// TIA Portal V20 export
FUNCTION_BLOCK "FB_LD_PressDemoAuto"   // FB, LAD
{ S7_Optimized_Access := 'TRUE' }
// stored: AutoNumber true
   VAR_INPUT
      Run { ExternalWritable := 'False'} : Bool;
      Reset { ExternalWritable := 'False'} : Bool;
      OwnerIndex { ExternalWritable := 'False'} : DInt;
      Delta { ExternalWritable := 'False'} : Time;
      TransferSettleTime { ExternalWritable := 'False'} : Time;
      PartQuality { ExternalWritable := 'False'} : Bool;
      RequireTwoHandStart { ExternalWritable := 'False'} : Bool;
      SourcePath { ExternalWritable := 'False'} : String[80];
      PartPresent { ExternalWritable := 'False'} : Bool;
      AirPressureOk { ExternalWritable := 'False'} : Bool;
      TwoHandHeld { ExternalWritable := 'False'} : Bool;
      StartPulse { ExternalWritable := 'False'} : Bool;
      PressSettleTime { ExternalWritable := 'False'} : Time;
   END_VAR
   VAR_IN_OUT
      PressRam { ExternalAccessible := 'False'; ExternalVisible := 'False'; ExternalWritable := 'False'} : "FB_CylinderCM";
      Door { ExternalAccessible := 'False'; ExternalVisible := 'False'; ExternalWritable := 'False'} : "FB_CylinderCM";
      PartSlide { ExternalAccessible := 'False'; ExternalVisible := 'False'; ExternalWritable := 'False'} : "FB_CylinderCM";
      Core { ExternalAccessible := 'False'; ExternalVisible := 'False'; ExternalWritable := 'False'} : "FRK_Core";
      Unit { ExternalAccessible := 'False'; ExternalVisible := 'False'; ExternalWritable := 'False'} : "FRK_Unit";
      Status { ExternalAccessible := 'False'; ExternalVisible := 'False'; ExternalWritable := 'False'} : "ST_ModuleStatus";
      Part { ExternalAccessible := 'False'; ExternalVisible := 'False'; ExternalWritable := 'False'} : "ST_PartContext";
      AlarmLog { ExternalAccessible := 'False'; ExternalVisible := 'False'; ExternalWritable := 'False'} : "FRK_AlarmLog";
   END_VAR
   VAR
      Seq { ExternalWritable := 'False'} : "FRK_SequenceCtx";
      Row1 { ExternalWritable := 'False'} : "FRK_SequenceRow";
      Row2 { ExternalWritable := 'False'} : "FRK_SequenceRow";
      Row3 { ExternalWritable := 'False'} : "FRK_SequenceRow";
      Row4 { ExternalWritable := 'False'} : "FRK_SequenceRow";
      Row5 { ExternalWritable := 'False'} : "FRK_SequenceRow";
      Row6 { ExternalWritable := 'False'} : "FRK_SequenceRow";
      Row7 { ExternalWritable := 'False'} : "FRK_SequenceRow";
      Row8 { ExternalWritable := 'False'} : "FRK_SequenceRow";
      Row9 { ExternalWritable := 'False'} : "FRK_SequenceRow";
      Row10 { ExternalWritable := 'False'} : "FRK_SequenceRow";
      Row11 { ExternalWritable := 'False'} : "FRK_SequenceRow";
      Row12 { ExternalWritable := 'False'} : "FRK_SequenceRow";
      Row13 { ExternalWritable := 'False'} : "FRK_SequenceRow";
      Row14 { ExternalWritable := 'False'} : "FRK_SequenceRow";
      Row15 { ExternalWritable := 'False'} : "FRK_SequenceRow";
      Row16 { ExternalWritable := 'False'} : "FRK_SequenceRow";
      At0 { ExternalAccessible := 'False'; ExternalVisible := 'False'; ExternalWritable := 'False'} : Bool;
      At100 { ExternalAccessible := 'False'; ExternalVisible := 'False'; ExternalWritable := 'False'} : Bool;
      At110 { ExternalAccessible := 'False'; ExternalVisible := 'False'; ExternalWritable := 'False'} : Bool;
      At130 { ExternalAccessible := 'False'; ExternalVisible := 'False'; ExternalWritable := 'False'} : Bool;
      At150 { ExternalAccessible := 'False'; ExternalVisible := 'False'; ExternalWritable := 'False'} : Bool;
      At170 { ExternalAccessible := 'False'; ExternalVisible := 'False'; ExternalWritable := 'False'} : Bool;
      At180 { ExternalAccessible := 'False'; ExternalVisible := 'False'; ExternalWritable := 'False'} : Bool;
      At185 { ExternalAccessible := 'False'; ExternalVisible := 'False'; ExternalWritable := 'False'} : Bool;
      At190 { ExternalAccessible := 'False'; ExternalVisible := 'False'; ExternalWritable := 'False'} : Bool;
      At200 { ExternalAccessible := 'False'; ExternalVisible := 'False'; ExternalWritable := 'False'} : Bool;
      At210 { ExternalAccessible := 'False'; ExternalVisible := 'False'; ExternalWritable := 'False'} : Bool;
      At215 { ExternalAccessible := 'False'; ExternalVisible := 'False'; ExternalWritable := 'False'} : Bool;
      At220 { ExternalAccessible := 'False'; ExternalVisible := 'False'; ExternalWritable := 'False'} : Bool;
      At230 { ExternalAccessible := 'False'; ExternalVisible := 'False'; ExternalWritable := 'False'} : Bool;
      At240 { ExternalAccessible := 'False'; ExternalVisible := 'False'; ExternalWritable := 'False'} : Bool;
      At999 { ExternalAccessible := 'False'; ExternalVisible := 'False'; ExternalWritable := 'False'} : Bool;
      Ready1 { ExternalAccessible := 'False'; ExternalVisible := 'False'; ExternalWritable := 'False'} : Bool;
      Ready2 { ExternalAccessible := 'False'; ExternalVisible := 'False'; ExternalWritable := 'False'} : Bool;
      Ready3 { ExternalAccessible := 'False'; ExternalVisible := 'False'; ExternalWritable := 'False'} : Bool;
      Ready4 { ExternalAccessible := 'False'; ExternalVisible := 'False'; ExternalWritable := 'False'} : Bool;
      Ready5 { ExternalAccessible := 'False'; ExternalVisible := 'False'; ExternalWritable := 'False'} : Bool;
      Advance { ExternalAccessible := 'False'; ExternalVisible := 'False'; ExternalWritable := 'False'} : Bool;
      Cycle { ExternalAccessible := 'False'; ExternalVisible := 'False'; ExternalWritable := 'False'} : "ST_PressDemoCycle";
      LoadPosition { ExternalAccessible := 'False'; ExternalVisible := 'False'; ExternalWritable := 'False'} : "FB_PressDemoLoadPosition";
      LoadDone { ExternalAccessible := 'False'; ExternalVisible := 'False'; ExternalWritable := 'False'} : Bool;
      LoadActive { ExternalAccessible := 'False'; ExternalVisible := 'False'; ExternalWritable := 'False'} : Bool;
   END_VAR
BEGIN

REGION Network 1
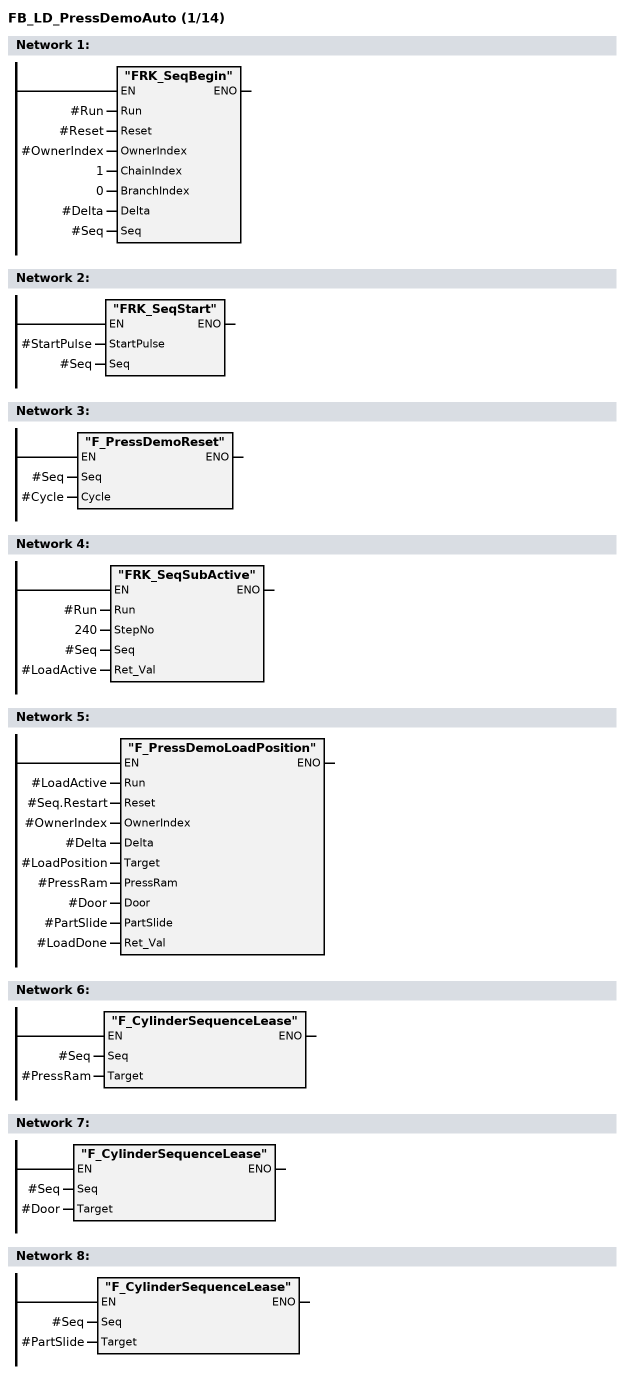
   RUNG wire#powerrail
      "FRK_SeqBegin"(Run := #Run, Reset := #Reset, OwnerIndex := #OwnerIndex, ChainIndex := 1, BranchIndex := 0, Delta := #Delta, Seq := #Seq)
   END_RUNG
   // the same network as SCL:
   "FRK_SeqBegin"(Run := #Run,
                  Reset := #Reset,
                  OwnerIndex := #OwnerIndex,
                  ChainIndex := 1,
                  BranchIndex := 0,
                  Delta := #Delta,
                  Seq := #Seq);
END_REGION

REGION Network 2
   RUNG wire#powerrail
      "FRK_SeqStart"(StartPulse := #StartPulse, Seq := #Seq)
   END_RUNG
   // the same network as SCL:
   "FRK_SeqStart"(StartPulse := #StartPulse, Seq := #Seq);
END_REGION

REGION Network 3
   RUNG wire#powerrail
      "F_PressDemoReset"(Seq := #Seq, Cycle := #Cycle)
   END_RUNG
   // the same network as SCL:
   "F_PressDemoReset"(Seq := #Seq, Cycle := #Cycle);
END_REGION

REGION Network 4
   RUNG wire#powerrail
      "FRK_SeqSubActive"(Run := #Run, StepNo := 240, Seq := #Seq, Ret_Val := #LoadActive)
   END_RUNG
   // the same network as SCL:
   "FRK_SeqSubActive"(Run := #Run, StepNo := 240, Seq := #Seq, Ret_Val := #LoadActive);
END_REGION

REGION Network 5
   RUNG wire#powerrail
      "F_PressDemoLoadPosition"(Run := #LoadActive, Reset := #Seq.Restart, OwnerIndex := #OwnerIndex, Delta := #Delta, Target := #LoadPosition, PressRam := #PressRam, Door := #Door, PartSlide := #PartSlide, Ret_Val := #LoadDone)
   END_RUNG
   // the same network as SCL:
   "F_PressDemoLoadPosition"(Run := #LoadActive,
                           Reset := #Seq.Restart,
                           OwnerIndex := #OwnerIndex,
                           Delta := #Delta,
                           Target := #LoadPosition,
                           PressRam := #PressRam,
                           Door := #Door,
                           PartSlide := #PartSlide,
                           Ret_Val := #LoadDone);
END_REGION

REGION Network 6
   RUNG wire#powerrail
      "F_CylinderSequenceLease"(Seq := #Seq, Target := #PressRam)
   END_RUNG
   // the same network as SCL:
   "F_CylinderSequenceLease"(Seq := #Seq, Target := #PressRam);
END_REGION

REGION Network 7
   RUNG wire#powerrail
      "F_CylinderSequenceLease"(Seq := #Seq, Target := #Door)
   END_RUNG
   // the same network as SCL:
   "F_CylinderSequenceLease"(Seq := #Seq, Target := #Door);
END_REGION

REGION Network 8
   RUNG wire#powerrail
      "F_CylinderSequenceLease"(Seq := #Seq, Target := #PartSlide)
   END_RUNG
   // the same network as SCL:
   "F_CylinderSequenceLease"(Seq := #Seq, Target := #PartSlide);
END_REGION

REGION Network 9
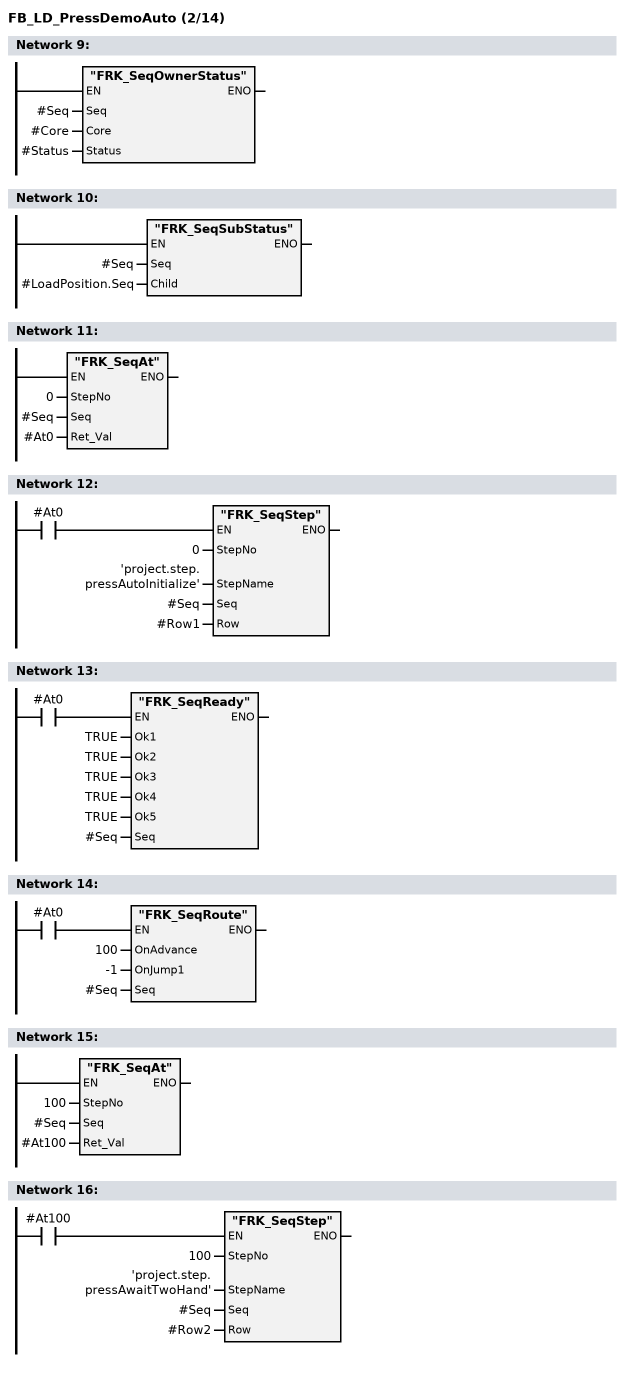
   RUNG wire#powerrail
      "FRK_SeqOwnerStatus"(Seq := #Seq, Core := #Core, Status := #Status)
   END_RUNG
   // the same network as SCL:
   "FRK_SeqOwnerStatus"(Seq := #Seq, Core := #Core, Status := #Status);
END_REGION

REGION Network 10
   RUNG wire#powerrail
      "FRK_SeqSubStatus"(Seq := #Seq, Child := #LoadPosition.Seq)
   END_RUNG
   // the same network as SCL:
   "FRK_SeqSubStatus"(Seq := #Seq, Child := #LoadPosition.Seq);
END_REGION

REGION Network 11
   RUNG wire#powerrail
      "FRK_SeqAt"(StepNo := 0, Seq := #Seq, Ret_Val := #At0)
   END_RUNG
   // the same network as SCL:
   "FRK_SeqAt"(StepNo := 0, Seq := #Seq, Ret_Val := #At0);
END_REGION

REGION Network 12
   IF #At0 THEN
       "FRK_SeqStep"(StepNo := 0, StepName := 'project.step.pressAutoInitialize', Seq := #Seq, Row := #Row1);
   END_IF;
END_REGION

REGION Network 13
   IF #At0 THEN
       "FRK_SeqReady"(Ok1 := TRUE, Ok2 := TRUE, Ok3 := TRUE, Ok4 := TRUE, Ok5 := TRUE, Seq := #Seq);
   END_IF;
END_REGION

REGION Network 14
   IF #At0 THEN "FRK_SeqRoute"(OnAdvance := 100, OnJump1 := -1, Seq := #Seq); END_IF;
END_REGION

REGION Network 15
   RUNG wire#powerrail
      "FRK_SeqAt"(StepNo := 100, Seq := #Seq, Ret_Val := #At100)
   END_RUNG
   // the same network as SCL:
   "FRK_SeqAt"(StepNo := 100, Seq := #Seq, Ret_Val := #At100);
END_REGION

REGION Network 16
   IF #At100 THEN
       "FRK_SeqStep"(StepNo := 100, StepName := 'project.step.pressAwaitTwoHand', Seq := #Seq, Row := #Row2);
   END_IF;
END_REGION

REGION Network 17
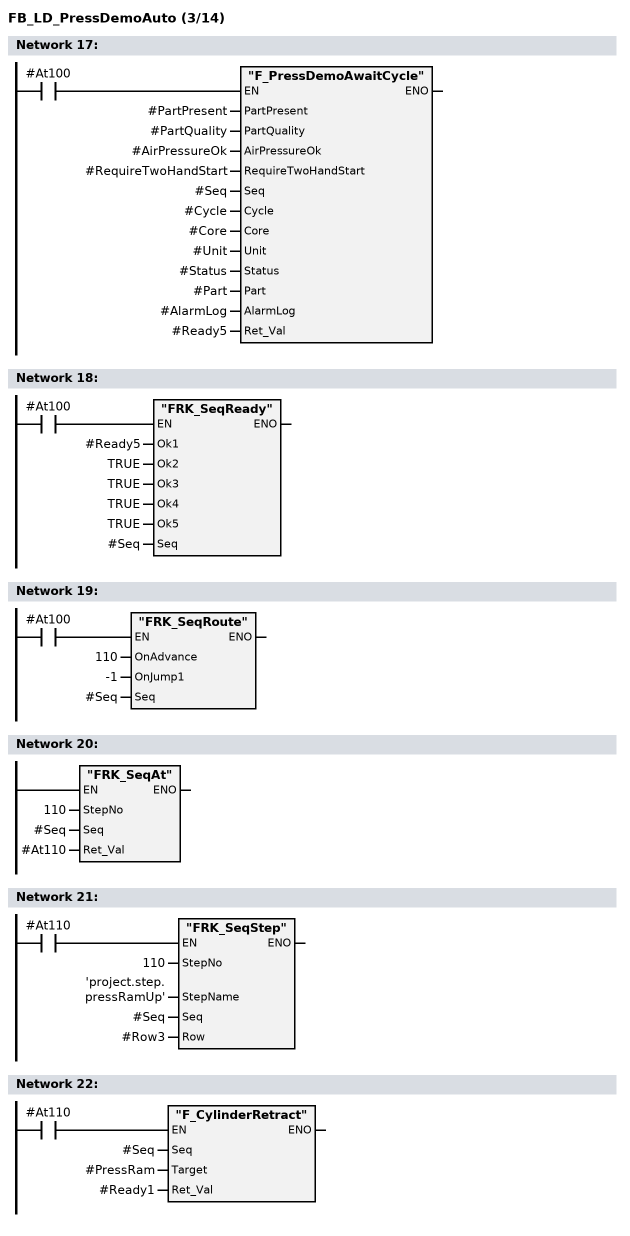
   IF #At100 THEN
       "F_PressDemoAwaitCycle"(PartPresent := #PartPresent,
                               PartQuality := #PartQuality,
                               AirPressureOk := #AirPressureOk,
                               RequireTwoHandStart := #RequireTwoHandStart,
                               Seq := #Seq,
                               Cycle := #Cycle,
                               Core := #Core,
                               Unit := #Unit,
                               Status := #Status,
                               Part := #Part,
                               AlarmLog := #AlarmLog,
                               Ret_Val := #Ready5);
   END_IF;
END_REGION

REGION Network 18
   IF #At100 THEN
       "FRK_SeqReady"(Ok1 := #Ready5, Ok2 := TRUE, Ok3 := TRUE, Ok4 := TRUE, Ok5 := TRUE, Seq := #Seq);
   END_IF;
END_REGION

REGION Network 19
   IF #At100 THEN "FRK_SeqRoute"(OnAdvance := 110, OnJump1 := -1, Seq := #Seq); END_IF;
END_REGION

REGION Network 20
   RUNG wire#powerrail
      "FRK_SeqAt"(StepNo := 110, Seq := #Seq, Ret_Val := #At110)
   END_RUNG
   // the same network as SCL:
   "FRK_SeqAt"(StepNo := 110, Seq := #Seq, Ret_Val := #At110);
END_REGION

REGION Network 21
   IF #At110 THEN
       "FRK_SeqStep"(StepNo := 110, StepName := 'project.step.pressRamUp', Seq := #Seq, Row := #Row3);
   END_IF;
END_REGION

REGION Network 22
   IF #At110 THEN "F_CylinderRetract"(Seq := #Seq, Target := #PressRam, Ret_Val := #Ready1); END_IF;
END_REGION

REGION Network 23
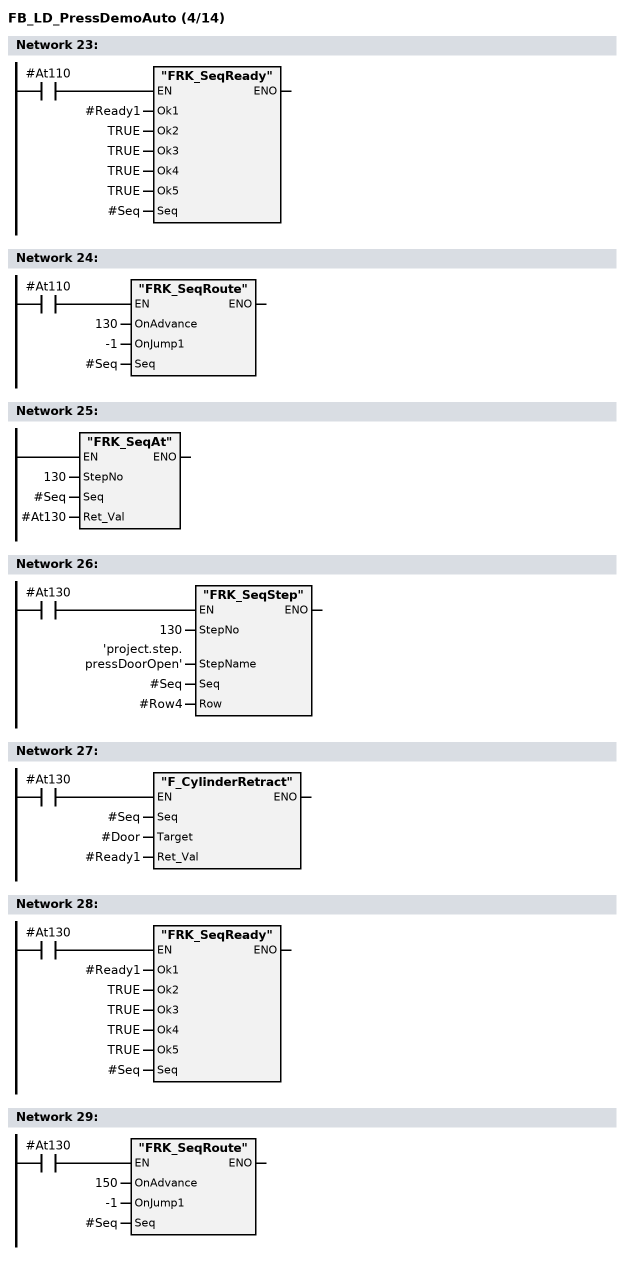
   IF #At110 THEN
       "FRK_SeqReady"(Ok1 := #Ready1, Ok2 := TRUE, Ok3 := TRUE, Ok4 := TRUE, Ok5 := TRUE, Seq := #Seq);
   END_IF;
END_REGION

REGION Network 24
   IF #At110 THEN "FRK_SeqRoute"(OnAdvance := 130, OnJump1 := -1, Seq := #Seq); END_IF;
END_REGION

REGION Network 25
   RUNG wire#powerrail
      "FRK_SeqAt"(StepNo := 130, Seq := #Seq, Ret_Val := #At130)
   END_RUNG
   // the same network as SCL:
   "FRK_SeqAt"(StepNo := 130, Seq := #Seq, Ret_Val := #At130);
END_REGION

REGION Network 26
   IF #At130 THEN
       "FRK_SeqStep"(StepNo := 130, StepName := 'project.step.pressDoorOpen', Seq := #Seq, Row := #Row4);
   END_IF;
END_REGION

REGION Network 27
   IF #At130 THEN "F_CylinderRetract"(Seq := #Seq, Target := #Door, Ret_Val := #Ready1); END_IF;
END_REGION

REGION Network 28
   IF #At130 THEN
       "FRK_SeqReady"(Ok1 := #Ready1, Ok2 := TRUE, Ok3 := TRUE, Ok4 := TRUE, Ok5 := TRUE, Seq := #Seq);
   END_IF;
END_REGION

REGION Network 29
   IF #At130 THEN "FRK_SeqRoute"(OnAdvance := 150, OnJump1 := -1, Seq := #Seq); END_IF;
END_REGION

REGION Network 30
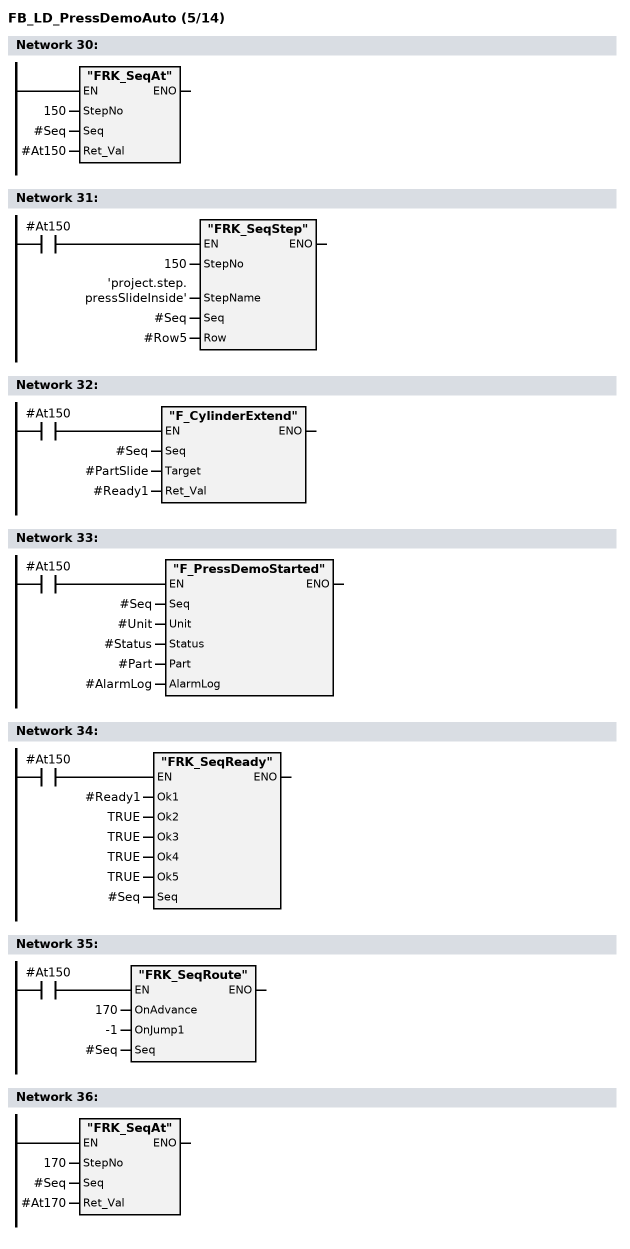
   RUNG wire#powerrail
      "FRK_SeqAt"(StepNo := 150, Seq := #Seq, Ret_Val := #At150)
   END_RUNG
   // the same network as SCL:
   "FRK_SeqAt"(StepNo := 150, Seq := #Seq, Ret_Val := #At150);
END_REGION

REGION Network 31
   IF #At150 THEN
       "FRK_SeqStep"(StepNo := 150, StepName := 'project.step.pressSlideInside', Seq := #Seq, Row := #Row5);
   END_IF;
END_REGION

REGION Network 32
   IF #At150 THEN "F_CylinderExtend"(Seq := #Seq, Target := #PartSlide, Ret_Val := #Ready1); END_IF;
END_REGION

REGION Network 33
   IF #At150 THEN
       "F_PressDemoStarted"(Seq := #Seq, Unit := #Unit, Status := #Status, Part := #Part, AlarmLog := #AlarmLog);
   END_IF;
END_REGION

REGION Network 34
   IF #At150 THEN
       "FRK_SeqReady"(Ok1 := #Ready1, Ok2 := TRUE, Ok3 := TRUE, Ok4 := TRUE, Ok5 := TRUE, Seq := #Seq);
   END_IF;
END_REGION

REGION Network 35
   IF #At150 THEN "FRK_SeqRoute"(OnAdvance := 170, OnJump1 := -1, Seq := #Seq); END_IF;
END_REGION

REGION Network 36
   RUNG wire#powerrail
      "FRK_SeqAt"(StepNo := 170, Seq := #Seq, Ret_Val := #At170)
   END_RUNG
   // the same network as SCL:
   "FRK_SeqAt"(StepNo := 170, Seq := #Seq, Ret_Val := #At170);
END_REGION

REGION Network 37
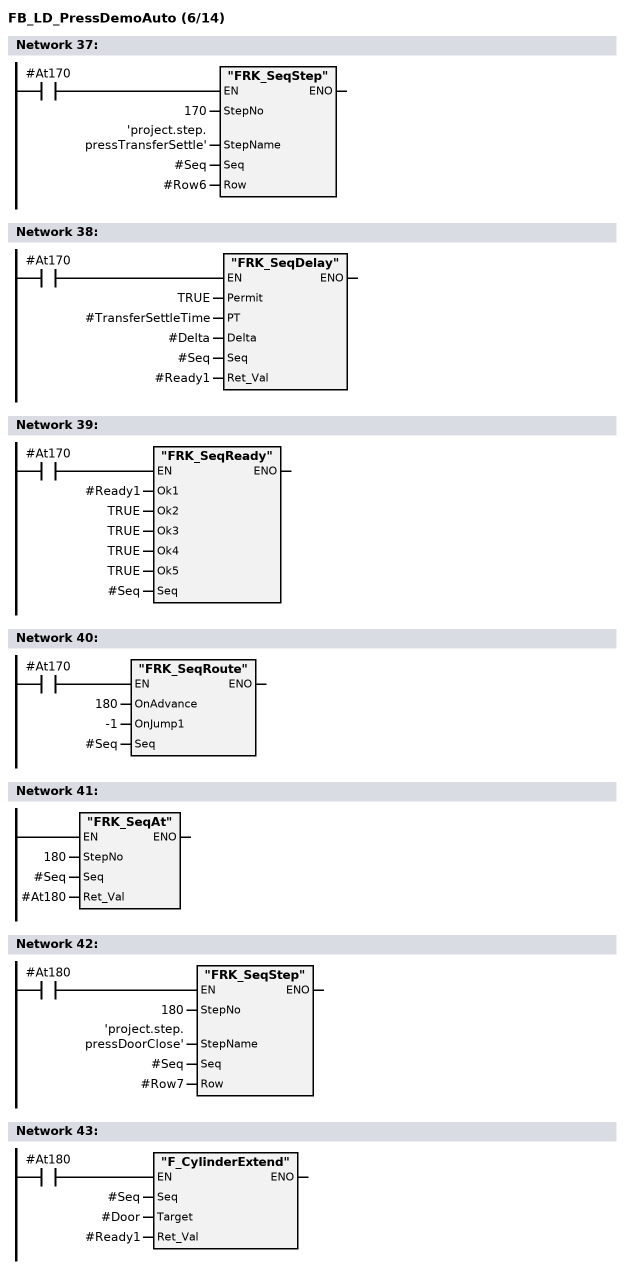
   IF #At170 THEN
       "FRK_SeqStep"(StepNo := 170, StepName := 'project.step.pressTransferSettle', Seq := #Seq, Row := #Row6);
   END_IF;
END_REGION

REGION Network 38
   IF #At170 THEN
       "FRK_SeqDelay"(Permit := TRUE, PT := #TransferSettleTime, Delta := #Delta, Seq := #Seq, Ret_Val := #Ready1);
   END_IF;
END_REGION

REGION Network 39
   IF #At170 THEN
       "FRK_SeqReady"(Ok1 := #Ready1, Ok2 := TRUE, Ok3 := TRUE, Ok4 := TRUE, Ok5 := TRUE, Seq := #Seq);
   END_IF;
END_REGION

REGION Network 40
   IF #At170 THEN "FRK_SeqRoute"(OnAdvance := 180, OnJump1 := -1, Seq := #Seq); END_IF;
END_REGION

REGION Network 41
   RUNG wire#powerrail
      "FRK_SeqAt"(StepNo := 180, Seq := #Seq, Ret_Val := #At180)
   END_RUNG
   // the same network as SCL:
   "FRK_SeqAt"(StepNo := 180, Seq := #Seq, Ret_Val := #At180);
END_REGION

REGION Network 42
   IF #At180 THEN
       "FRK_SeqStep"(StepNo := 180, StepName := 'project.step.pressDoorClose', Seq := #Seq, Row := #Row7);
   END_IF;
END_REGION

REGION Network 43
   IF #At180 THEN "F_CylinderExtend"(Seq := #Seq, Target := #Door, Ret_Val := #Ready1); END_IF;
END_REGION

REGION Network 44
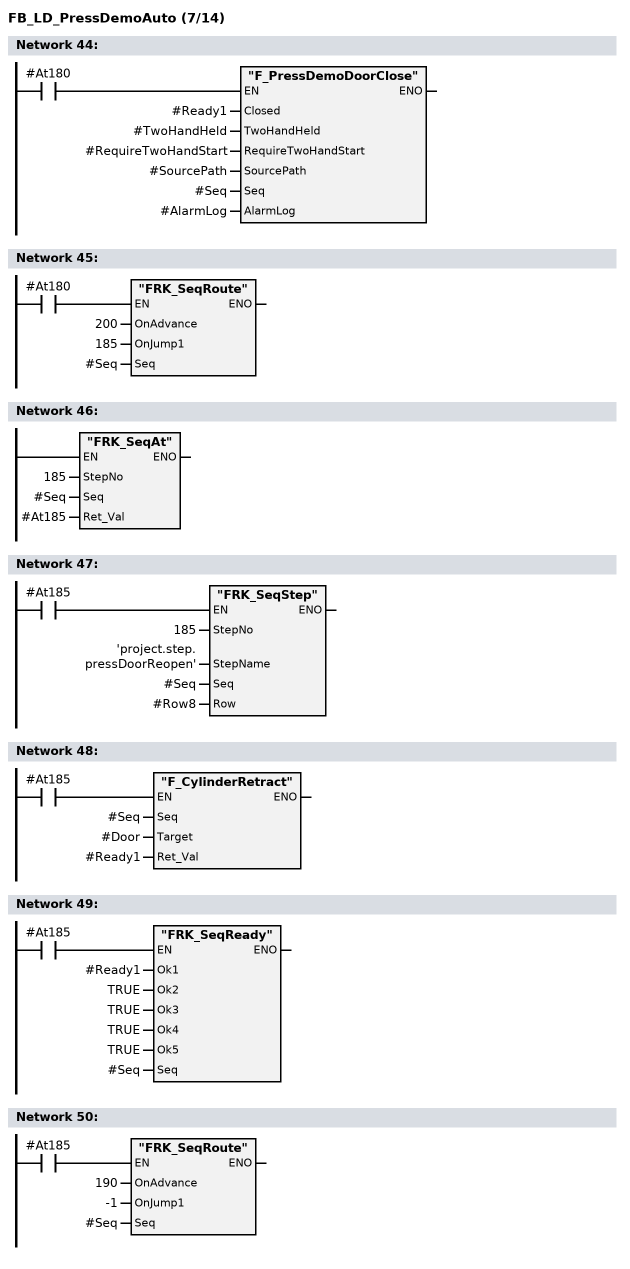
   IF #At180 THEN
       "F_PressDemoDoorClose"(Closed := #Ready1,
                              TwoHandHeld := #TwoHandHeld,
                              RequireTwoHandStart := #RequireTwoHandStart,
                              SourcePath := #SourcePath,
                              Seq := #Seq,
                              AlarmLog := #AlarmLog);
   END_IF;
END_REGION

REGION Network 45
   IF #At180 THEN "FRK_SeqRoute"(OnAdvance := 200, OnJump1 := 185, Seq := #Seq); END_IF;
END_REGION

REGION Network 46
   RUNG wire#powerrail
      "FRK_SeqAt"(StepNo := 185, Seq := #Seq, Ret_Val := #At185)
   END_RUNG
   // the same network as SCL:
   "FRK_SeqAt"(StepNo := 185, Seq := #Seq, Ret_Val := #At185);
END_REGION

REGION Network 47
   IF #At185 THEN
       "FRK_SeqStep"(StepNo := 185, StepName := 'project.step.pressDoorReopen', Seq := #Seq, Row := #Row8);
   END_IF;
END_REGION

REGION Network 48
   IF #At185 THEN "F_CylinderRetract"(Seq := #Seq, Target := #Door, Ret_Val := #Ready1); END_IF;
END_REGION

REGION Network 49
   IF #At185 THEN
       "FRK_SeqReady"(Ok1 := #Ready1, Ok2 := TRUE, Ok3 := TRUE, Ok4 := TRUE, Ok5 := TRUE, Seq := #Seq);
   END_IF;
END_REGION

REGION Network 50
   IF #At185 THEN "FRK_SeqRoute"(OnAdvance := 190, OnJump1 := -1, Seq := #Seq); END_IF;
END_REGION

REGION Network 51
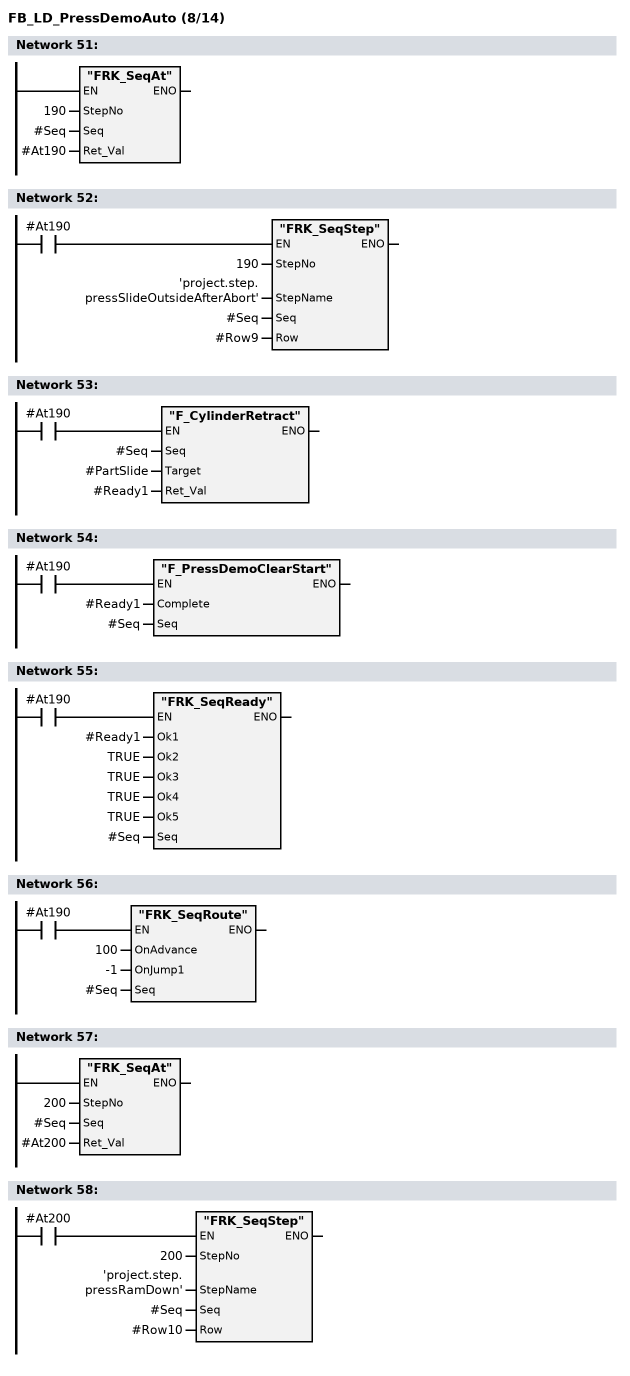
   RUNG wire#powerrail
      "FRK_SeqAt"(StepNo := 190, Seq := #Seq, Ret_Val := #At190)
   END_RUNG
   // the same network as SCL:
   "FRK_SeqAt"(StepNo := 190, Seq := #Seq, Ret_Val := #At190);
END_REGION

REGION Network 52
   IF #At190 THEN
       "FRK_SeqStep"(StepNo := 190,
                     StepName := 'project.step.pressSlideOutsideAfterAbort',
                     Seq := #Seq,
                     Row := #Row9);
   END_IF;
END_REGION

REGION Network 53
   IF #At190 THEN "F_CylinderRetract"(Seq := #Seq, Target := #PartSlide, Ret_Val := #Ready1); END_IF;
END_REGION

REGION Network 54
   IF #At190 THEN "F_PressDemoClearStart"(Complete := #Ready1, Seq := #Seq); END_IF;
END_REGION

REGION Network 55
   IF #At190 THEN
       "FRK_SeqReady"(Ok1 := #Ready1, Ok2 := TRUE, Ok3 := TRUE, Ok4 := TRUE, Ok5 := TRUE, Seq := #Seq);
   END_IF;
END_REGION

REGION Network 56
   IF #At190 THEN "FRK_SeqRoute"(OnAdvance := 100, OnJump1 := -1, Seq := #Seq); END_IF;
END_REGION

REGION Network 57
   RUNG wire#powerrail
      "FRK_SeqAt"(StepNo := 200, Seq := #Seq, Ret_Val := #At200)
   END_RUNG
   // the same network as SCL:
   "FRK_SeqAt"(StepNo := 200, Seq := #Seq, Ret_Val := #At200);
END_REGION

REGION Network 58
   IF #At200 THEN
       "FRK_SeqStep"(StepNo := 200, StepName := 'project.step.pressRamDown', Seq := #Seq, Row := #Row10);
   END_IF;
END_REGION

REGION Network 59
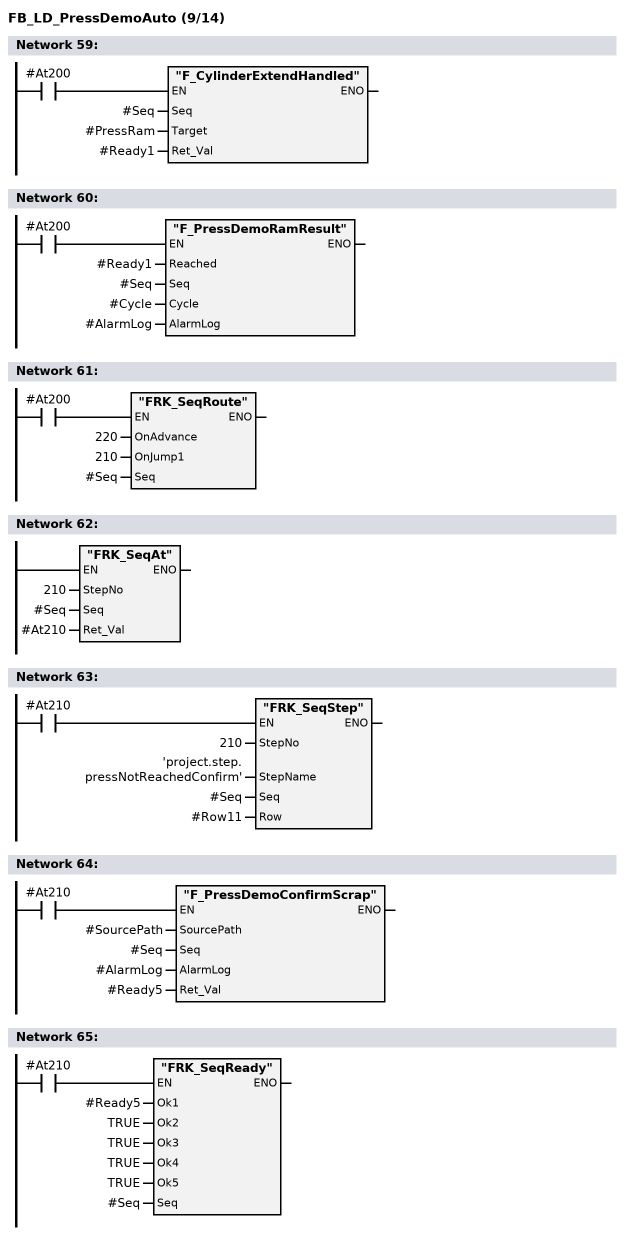
   IF #At200 THEN "F_CylinderExtendHandled"(Seq := #Seq, Target := #PressRam, Ret_Val := #Ready1); END_IF;
END_REGION

REGION Network 60
   IF #At200 THEN
       "F_PressDemoRamResult"(Reached := #Ready1, Seq := #Seq, Cycle := #Cycle, AlarmLog := #AlarmLog);
   END_IF;
END_REGION

REGION Network 61
   IF #At200 THEN "FRK_SeqRoute"(OnAdvance := 220, OnJump1 := 210, Seq := #Seq); END_IF;
END_REGION

REGION Network 62
   RUNG wire#powerrail
      "FRK_SeqAt"(StepNo := 210, Seq := #Seq, Ret_Val := #At210)
   END_RUNG
   // the same network as SCL:
   "FRK_SeqAt"(StepNo := 210, Seq := #Seq, Ret_Val := #At210);
END_REGION

REGION Network 63
   IF #At210 THEN
       "FRK_SeqStep"(StepNo := 210, StepName := 'project.step.pressNotReachedConfirm', Seq := #Seq, Row := #Row11);
   END_IF;
END_REGION

REGION Network 64
   IF #At210 THEN
       "F_PressDemoConfirmScrap"(SourcePath := #SourcePath, Seq := #Seq, AlarmLog := #AlarmLog, Ret_Val := #Ready5);
   END_IF;
END_REGION

REGION Network 65
   IF #At210 THEN
       "FRK_SeqReady"(Ok1 := #Ready5, Ok2 := TRUE, Ok3 := TRUE, Ok4 := TRUE, Ok5 := TRUE, Seq := #Seq);
   END_IF;
END_REGION

REGION Network 66
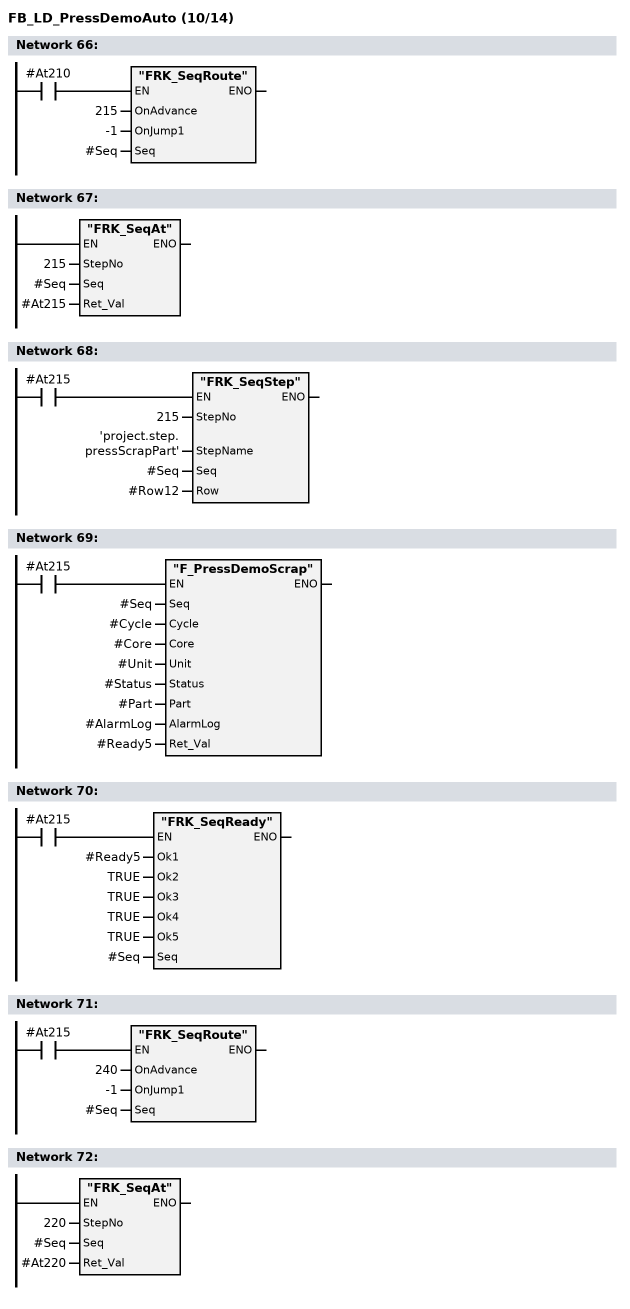
   IF #At210 THEN "FRK_SeqRoute"(OnAdvance := 215, OnJump1 := -1, Seq := #Seq); END_IF;
END_REGION

REGION Network 67
   RUNG wire#powerrail
      "FRK_SeqAt"(StepNo := 215, Seq := #Seq, Ret_Val := #At215)
   END_RUNG
   // the same network as SCL:
   "FRK_SeqAt"(StepNo := 215, Seq := #Seq, Ret_Val := #At215);
END_REGION

REGION Network 68
   IF #At215 THEN
       "FRK_SeqStep"(StepNo := 215, StepName := 'project.step.pressScrapPart', Seq := #Seq, Row := #Row12);
   END_IF;
END_REGION

REGION Network 69
   IF #At215 THEN
       "F_PressDemoScrap"(Seq := #Seq,
                          Cycle := #Cycle,
                          Core := #Core,
                          Unit := #Unit,
                          Status := #Status,
                          Part := #Part,
                          AlarmLog := #AlarmLog,
                          Ret_Val := #Ready5);
   END_IF;
END_REGION

REGION Network 70
   IF #At215 THEN
       "FRK_SeqReady"(Ok1 := #Ready5, Ok2 := TRUE, Ok3 := TRUE, Ok4 := TRUE, Ok5 := TRUE, Seq := #Seq);
   END_IF;
END_REGION

REGION Network 71
   IF #At215 THEN "FRK_SeqRoute"(OnAdvance := 240, OnJump1 := -1, Seq := #Seq); END_IF;
END_REGION

REGION Network 72
   RUNG wire#powerrail
      "FRK_SeqAt"(StepNo := 220, Seq := #Seq, Ret_Val := #At220)
   END_RUNG
   // the same network as SCL:
   "FRK_SeqAt"(StepNo := 220, Seq := #Seq, Ret_Val := #At220);
END_REGION

REGION Network 73
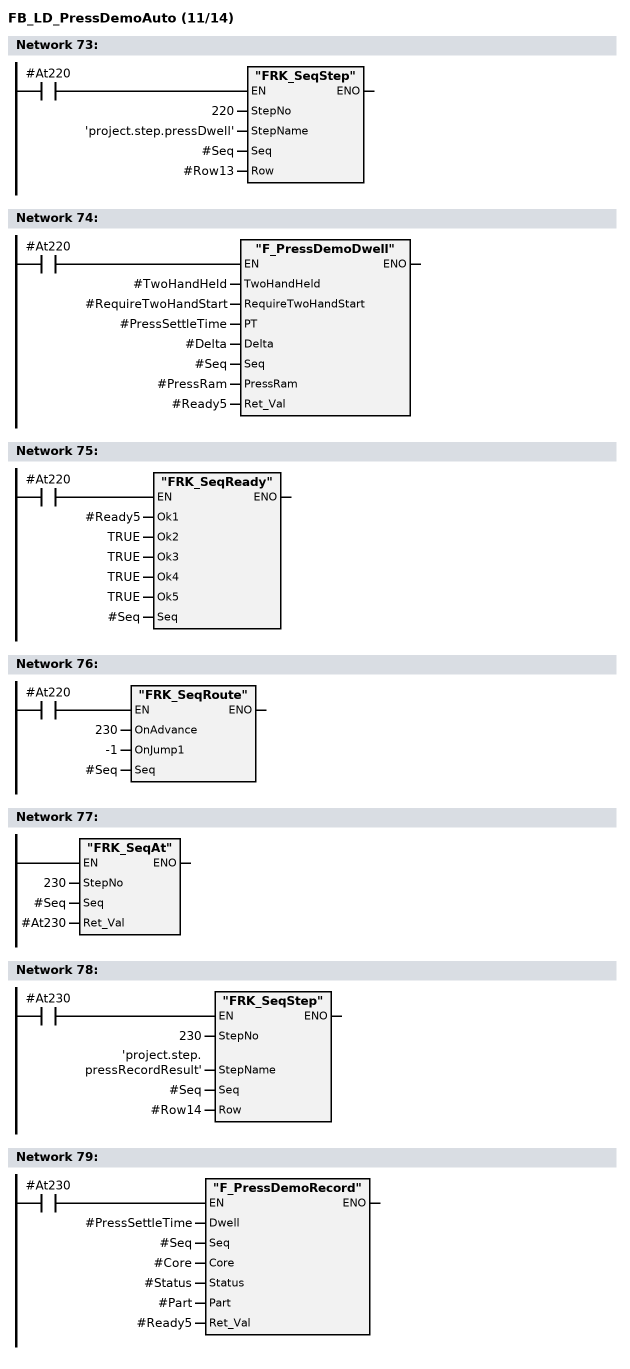
   IF #At220 THEN
       "FRK_SeqStep"(StepNo := 220, StepName := 'project.step.pressDwell', Seq := #Seq, Row := #Row13);
   END_IF;
END_REGION

REGION Network 74
   IF #At220 THEN
       "F_PressDemoDwell"(TwoHandHeld := #TwoHandHeld,
                          RequireTwoHandStart := #RequireTwoHandStart,
                          PT := #PressSettleTime,
                          Delta := #Delta,
                          Seq := #Seq,
                          PressRam := #PressRam,
                          Ret_Val := #Ready5);
   END_IF;
END_REGION

REGION Network 75
   IF #At220 THEN
       "FRK_SeqReady"(Ok1 := #Ready5, Ok2 := TRUE, Ok3 := TRUE, Ok4 := TRUE, Ok5 := TRUE, Seq := #Seq);
   END_IF;
END_REGION

REGION Network 76
   IF #At220 THEN "FRK_SeqRoute"(OnAdvance := 230, OnJump1 := -1, Seq := #Seq); END_IF;
END_REGION

REGION Network 77
   RUNG wire#powerrail
      "FRK_SeqAt"(StepNo := 230, Seq := #Seq, Ret_Val := #At230)
   END_RUNG
   // the same network as SCL:
   "FRK_SeqAt"(StepNo := 230, Seq := #Seq, Ret_Val := #At230);
END_REGION

REGION Network 78
   IF #At230 THEN
       "FRK_SeqStep"(StepNo := 230, StepName := 'project.step.pressRecordResult', Seq := #Seq, Row := #Row14);
   END_IF;
END_REGION

REGION Network 79
   IF #At230 THEN
       "F_PressDemoRecord"(Dwell := #PressSettleTime,
                           Seq := #Seq,
                           Core := #Core,
                           Status := #Status,
                           Part := #Part,
                           Ret_Val := #Ready5);
   END_IF;
END_REGION

REGION Network 80
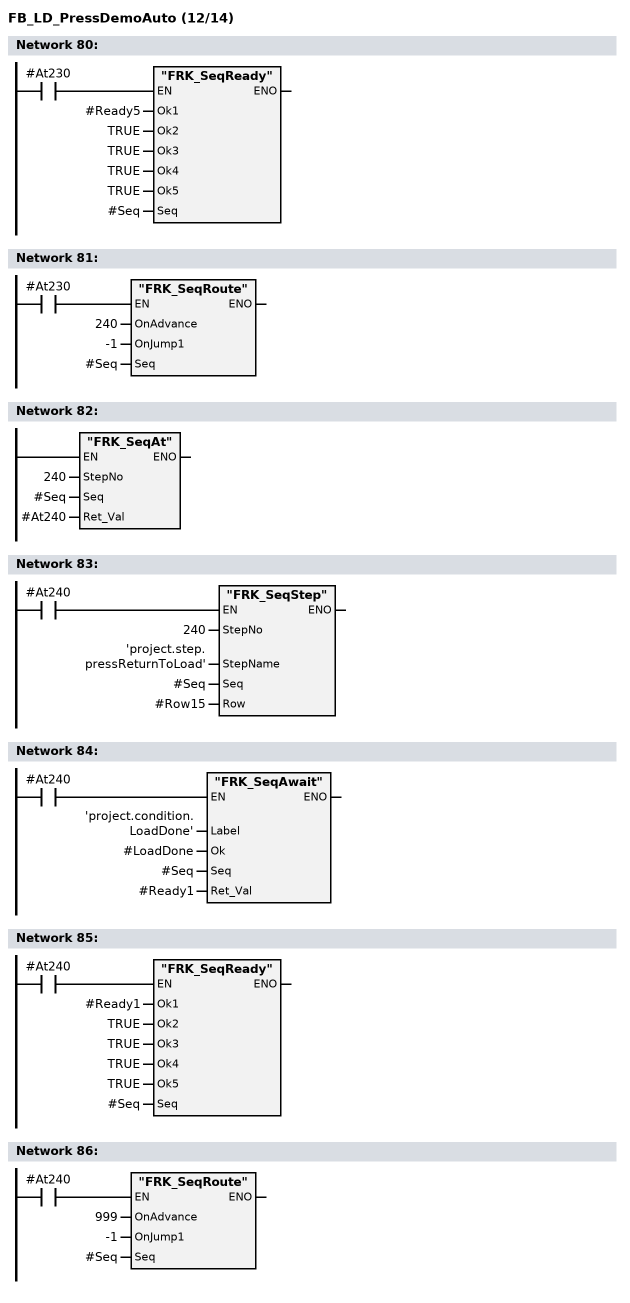
   IF #At230 THEN
       "FRK_SeqReady"(Ok1 := #Ready5, Ok2 := TRUE, Ok3 := TRUE, Ok4 := TRUE, Ok5 := TRUE, Seq := #Seq);
   END_IF;
END_REGION

REGION Network 81
   IF #At230 THEN "FRK_SeqRoute"(OnAdvance := 240, OnJump1 := -1, Seq := #Seq); END_IF;
END_REGION

REGION Network 82
   RUNG wire#powerrail
      "FRK_SeqAt"(StepNo := 240, Seq := #Seq, Ret_Val := #At240)
   END_RUNG
   // the same network as SCL:
   "FRK_SeqAt"(StepNo := 240, Seq := #Seq, Ret_Val := #At240);
END_REGION

REGION Network 83
   IF #At240 THEN
       "FRK_SeqStep"(StepNo := 240, StepName := 'project.step.pressReturnToLoad', Seq := #Seq, Row := #Row15);
   END_IF;
END_REGION

REGION Network 84
   IF #At240 THEN
       "FRK_SeqAwait"(Label := 'project.condition.LoadDone', Ok := #LoadDone, Seq := #Seq, Ret_Val := #Ready1);
   END_IF;
END_REGION

REGION Network 85
   IF #At240 THEN
       "FRK_SeqReady"(Ok1 := #Ready1, Ok2 := TRUE, Ok3 := TRUE, Ok4 := TRUE, Ok5 := TRUE, Seq := #Seq);
   END_IF;
END_REGION

REGION Network 86
   IF #At240 THEN "FRK_SeqRoute"(OnAdvance := 999, OnJump1 := -1, Seq := #Seq); END_IF;
END_REGION

REGION Network 87
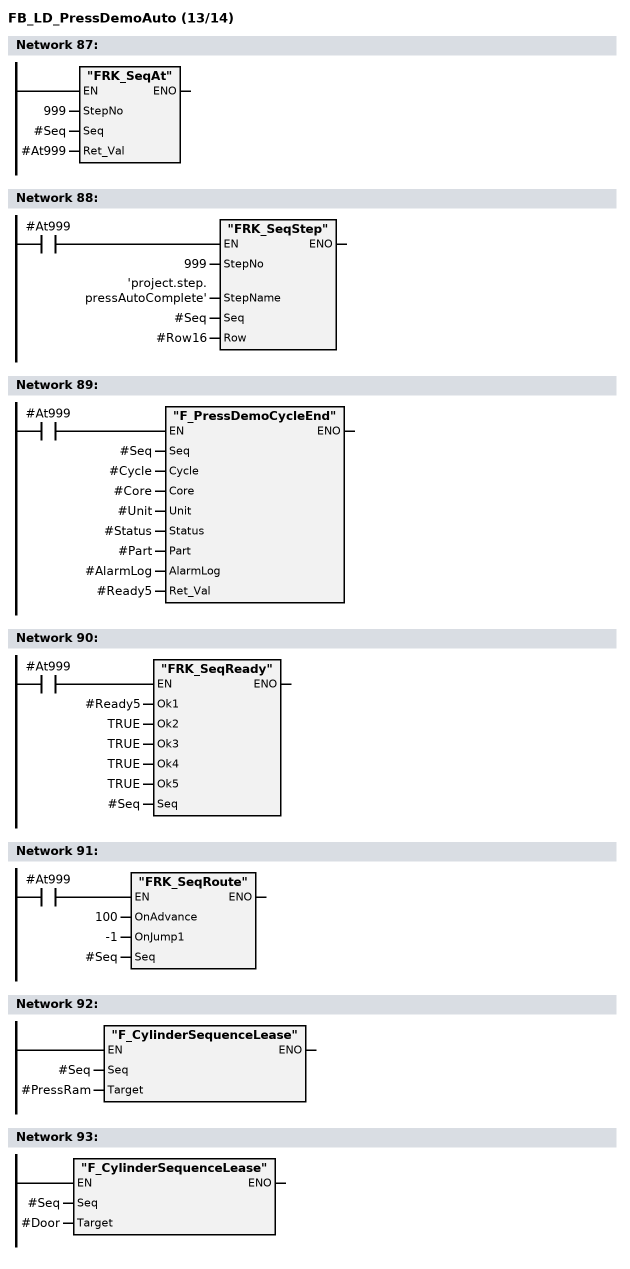
   RUNG wire#powerrail
      "FRK_SeqAt"(StepNo := 999, Seq := #Seq, Ret_Val := #At999)
   END_RUNG
   // the same network as SCL:
   "FRK_SeqAt"(StepNo := 999, Seq := #Seq, Ret_Val := #At999);
END_REGION

REGION Network 88
   IF #At999 THEN
       "FRK_SeqStep"(StepNo := 999, StepName := 'project.step.pressAutoComplete', Seq := #Seq, Row := #Row16);
   END_IF;
END_REGION

REGION Network 89
   IF #At999 THEN
       "F_PressDemoCycleEnd"(Seq := #Seq,
                             Cycle := #Cycle,
                             Core := #Core,
                             Unit := #Unit,
                             Status := #Status,
                             Part := #Part,
                             AlarmLog := #AlarmLog,
                             Ret_Val := #Ready5);
   END_IF;
END_REGION

REGION Network 90
   IF #At999 THEN
       "FRK_SeqReady"(Ok1 := #Ready5, Ok2 := TRUE, Ok3 := TRUE, Ok4 := TRUE, Ok5 := TRUE, Seq := #Seq);
   END_IF;
END_REGION

REGION Network 91
   IF #At999 THEN "FRK_SeqRoute"(OnAdvance := 100, OnJump1 := -1, Seq := #Seq); END_IF;
END_REGION

REGION Network 92
   RUNG wire#powerrail
      "F_CylinderSequenceLease"(Seq := #Seq, Target := #PressRam)
   END_RUNG
   // the same network as SCL:
   "F_CylinderSequenceLease"(Seq := #Seq, Target := #PressRam);
END_REGION

REGION Network 93
   RUNG wire#powerrail
      "F_CylinderSequenceLease"(Seq := #Seq, Target := #Door)
   END_RUNG
   // the same network as SCL:
   "F_CylinderSequenceLease"(Seq := #Seq, Target := #Door);
END_REGION

REGION Network 94
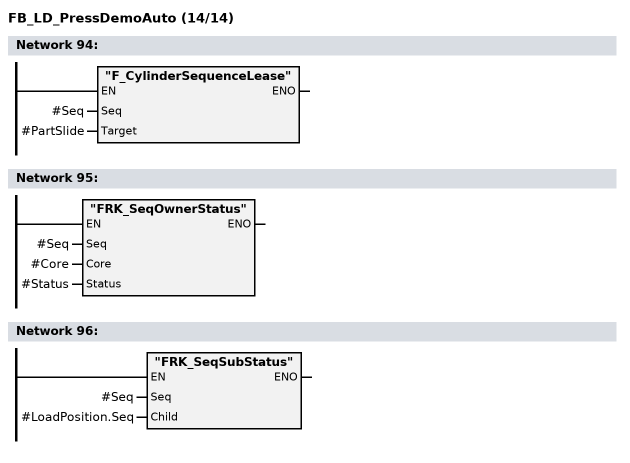
   RUNG wire#powerrail
      "F_CylinderSequenceLease"(Seq := #Seq, Target := #PartSlide)
   END_RUNG
   // the same network as SCL:
   "F_CylinderSequenceLease"(Seq := #Seq, Target := #PartSlide);
END_REGION

REGION Network 95
   RUNG wire#powerrail
      "FRK_SeqOwnerStatus"(Seq := #Seq, Core := #Core, Status := #Status)
   END_RUNG
   // the same network as SCL:
   "FRK_SeqOwnerStatus"(Seq := #Seq, Core := #Core, Status := #Status);
END_REGION

REGION Network 96
   RUNG wire#powerrail
      "FRK_SeqSubStatus"(Seq := #Seq, Child := #LoadPosition.Seq)
   END_RUNG
   // the same network as SCL:
   "FRK_SeqSubStatus"(Seq := #Seq, Child := #LoadPosition.Seq);
END_REGION
END_FUNCTION_BLOCK
